// TIA Portal V20 export
// export: Created 2026-10-20T12:52:35.7624926Z, ExportSetting WithDefaults, DisplayName Totally Integrated Automation Portal, DisplayVersion V20 Update 6, DisplayName TIA Portal Openness, DisplayVersion V20 Update 6, DisplayName TIA Portal Version Control Interface, DisplayVersion V20 Update 6, DisplayName SINAMICS Startdrive Advanced, DisplayVersion V20 SP1, DisplayName SINAMICS Startdrive G130, G150, S120, S150, SINAMICS MV, G220, S200, S210, DisplayVersion V20 SP1, DisplayName SINAMICS Startdrive G110M, G120, G120C, G120D, G120P, G115D, DisplayVersion V20 SP1, DisplayName STEP 7 Professional, DisplayVersion V20 Update 6, DisplayName STEP 7 Safety, DisplayVersion V20 Update 2, DisplayName WinCC Basic/Comfort/Advanced, DisplayVersion V20 Update 6, DisplayName WinCC Unified, DisplayVersion V20 Update 6
FUNCTION "Pre_Safe" : Void   // FC1000, LAD
{ S7_Optimized_Access := 'TRUE' }
VERSION : 0.1
// stored: AutoNumber false, IsIECCheckEnabled false, SetENOAutomatically false, UDAEnableTagReadback false
BEGIN

REGION Network 1
   // "Receive_Data_from_LGX".RCV_LENGTH
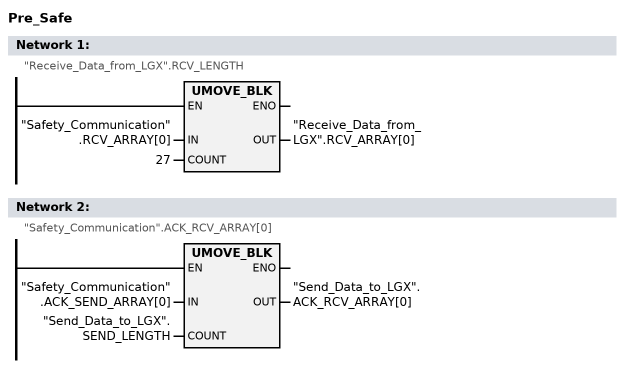
   UMOVE_BLK(IN := "Safety_Communication".RCV_ARRAY[0],
             COUNT := 27,
             OUT => "Receive_Data_from_LGX".RCV_ARRAY[0]);
END_REGION

REGION Network 2
   // "Safety_Communication".ACK_RCV_ARRAY[0]
   UMOVE_BLK(IN := "Safety_Communication".ACK_SEND_ARRAY[0],
             COUNT := "Send_Data_to_LGX".SEND_LENGTH,
             OUT => "Send_Data_to_LGX".ACK_RCV_ARRAY[0]);
END_REGION
END_FUNCTION
